TYPE "DT_MEASUREMENT_SYSTEM_CONTROL"
VERSION : 0.1
   STRUCT
      P { S7_SetPoint := 'False'} : "DT_MEASUREMENT_SOLO" := ((), (), FALSE, 1, 0, 168, 32000, 32000, 32000, 0, 0, 0, 0, 0, 0, 0, 0, 0, 0, 0, 0, 0, 0.0, 'kW');
      Q { S7_SetPoint := 'False'} : "DT_MEASUREMENT_SOLO" := ((), (), FALSE, 1, 0, 169, 32000, 32000, 32000, 0, 0, 0, 0, 0, 0, 0, 0, 0, 0, 0, 0, 0, 0.0, 'kVAr');
      S { S7_SetPoint := 'False'} : "DT_MEASUREMENT_SOLO" := ((), (), FALSE, 1, 0, 170, 32000, 32000, 32000, 0, 0, 0, 0, 0, 0, 0, 0, 0, 0, 0, 0, 0, 0.0, 'kVA');
      U_LL { S7_SetPoint := 'False'} : "DT_MEASUREMENT_SOLO" := ((), (), FALSE, 1, 0, 171, 32000, 32000, 32000, 0, 0, 0, 0, 0, 0, 0, 0, 0, 0, 0, 0, 0, 0.0, 'V');
      I { S7_SetPoint := 'False'} : "DT_MEASUREMENT_SOLO" := ((), (), FALSE, 1, 0, 172, 32000, 32000, 32000, 0, 0, 0, 0, 0, 0, 0, 0, 0, 0, 0, 0, 0, 0.0, 'A');
      PF { S7_SetPoint := 'False'} : "DT_MEASUREMENT_SOLO" := ((), (), FALSE, 1, 0, 173, 32000, 32000, 32000, 0, 0, 0, 0, 0, 0, 0, 0, 0, 0, 0, 0, 0, 0.0, '-');
      f_GEN { S7_SetPoint := 'False'} : "DT_MEASUREMENT_SOLO" := ((), (), FALSE, 1, 0, 174, 32000, 32000, 32000, 0, 0, 0, 0, 0, 0, 0, 0, 0, 0, 0, 0, 0, 0.0, 'Hz');
      f_GRID { S7_SetPoint := 'False'} : "DT_MEASUREMENT_SOLO" := ((), (), FALSE, 0, 0, 175, 32000, 32000, 32000, 0, 0, 0, 0, 0, 0, 0, 0, 0, 0, 0, 0, 0, 0.0, 'Hz');
      h { S7_SetPoint := 'False'} : "DT_MEASUREMENT_SOLO" := ((), (), FALSE, 1, 0, 176, 32000, 32000, 32000, 0, 0, 0, 0, 0, 0, 0, 0, 0, 0, 0, 0, 0, 0.0, 'm');
      pt { S7_SetPoint := 'False'} : "DT_MEASUREMENT_SOLO" := ((), (), FALSE, 1, 0, 177, 32000, 32000, 32000, 0, 0, 0, 0, 0, 0, 0, 0, 0, 0, 0, 0, 0, 0.0, 'bar');
      n { S7_SetPoint := 'False'} : "DT_MEASUREMENT_SOLO" := ((), (), FALSE, 1, 0, 178, 32000, 32000, 32000, 0, 0, 0, 0, 0, 0, 0, 0, 0, 0, 0, 0, 0, 0.0, 'rpm');
      MEAS_11 { S7_SetPoint := 'False'} : "DT_MEASUREMENT_SOLO" := ((), (), FALSE, 1, 0, 179, 32000, 32000, 32000, 0, 0, 0, 0, 0, 0, 0, 0, 0, 0, 0, 0, 0, 0.0, '');
      MEAS_12 { S7_SetPoint := 'False'} : "DT_MEASUREMENT_SOLO" := ((), (), FALSE, 1, 0, 180, 32000, 32000, 32000, 0, 0, 0, 0, 0, 0, 0, 0, 0, 0, 0, 0, 0, 0.0, '');
      MEAS_13 { S7_SetPoint := 'False'} : "DT_MEASUREMENT_SOLO" := ((), (), FALSE, 1, 0, 181, 32000, 32000, 32000, 0, 0, 0, 0, 0, 0, 0, 0, 0, 0, 0, 0, 0, 0.0, '');
      MEAS_14 { S7_SetPoint := 'False'} : "DT_MEASUREMENT_SOLO" := ((), (), FALSE, 1, 0, 182, 32000, 32000, 32000, 0, 0, 0, 0, 0, 0, 0, 0, 0, 0, 0, 0, 0, 0.0, '');
      MEAS_15 { S7_SetPoint := 'False'} : "DT_MEASUREMENT_SOLO" := ((), (), FALSE, 1, 0, 183, 32000, 32000, 32000, 0, 0, 0, 0, 0, 0, 0, 0, 0, 0, 0, 0, 0, 0.0, '');
      MEAS_16 { S7_SetPoint := 'False'} : "DT_MEASUREMENT_SOLO" := ((), (), FALSE, 1, 0, 184, 32000, 32000, 32000, 0, 0, 0, 0, 0, 0, 0, 0, 0, 0, 0, 0, 0, 0.0, '');
      MEAS_17 { S7_SetPoint := 'False'} : "DT_MEASUREMENT_SOLO" := ((), (), FALSE, 1, 0, 185, 32000, 32000, 32000, 0, 0, 0, 0, 0, 0, 0, 0, 0, 0, 0, 0, 0, 0.0, '');
      MEAS_18 { S7_SetPoint := 'False'} : "DT_MEASUREMENT_SOLO" := ((), (), FALSE, 1, 0, 186, 32000, 32000, 32000, 0, 0, 0, 0, 0, 0, 0, 0, 0, 0, 0, 0, 0, 0.0, '');
      MEAS_19 { S7_SetPoint := 'False'} : "DT_MEASUREMENT_SOLO" := ((), (), FALSE, 1, 0, 187, 32000, 32000, 32000, 0, 0, 0, 0, 0, 0, 0, 0, 0, 0, 0, 0, 0, 0.0, '');
      MEAS_20 { S7_SetPoint := 'False'} : "DT_MEASUREMENT_SOLO" := ((), (), FALSE, 1, 0, 188, 32000, 32000, 32000, 0, 0, 0, 0, 0, 0, 0, 0, 0, 0, 0, 0, 0, 0.0, '');
      MEAS_21 { S7_SetPoint := 'False'} : "DT_MEASUREMENT_SOLO" := ((), (), FALSE, 1, 0, 189, 32000, 32000, 32000, 0, 0, 0, 0, 0, 0, 0, 0, 0, 0, 0, 0, 0, 0.0, '');
      MEAS_22 { S7_SetPoint := 'False'} : "DT_MEASUREMENT_SOLO" := ((), (), FALSE, 1, 0, 190, 32000, 32000, 32000, 0, 0, 0, 0, 0, 0, 0, 0, 0, 0, 0, 0, 0, 0.0, '');
      MEAS_23 { S7_SetPoint := 'False'} : "DT_MEASUREMENT_SOLO" := ((), (), FALSE, 1, 0, 191, 32000, 32000, 32000, 0, 0, 0, 0, 0, 0, 0, 0, 0, 0, 0, 0, 0, 0.0, '');
   END_STRUCT;

END_TYPE

